(* IEC 61131-3 sources: MongoMation/docs, 1 file *)

(* ---- probe-sorting-by-height-basic.st ---- *)
(* I/O probe for scene sorting-by-height-basic (Sorting by Height (Basic)). Generated by scripts/gen-probe.ts. *)
PROGRAM io_probe
  VAR
    I0 AT %QX12.4 : BOOL; (* High sensor *)
    I1 AT %QX12.5 : BOOL; (* Low sensor *)
    I2 AT %QX12.6 : BOOL; (* Pallet sensor *)
    I3 AT %QX12.7 : BOOL; (* Loaded *)
    I4 AT %QX13.0 : BOOL; (* At left entry *)
    I5 AT %QX13.1 : BOOL; (* At left exit *)
    I6 AT %QX13.2 : BOOL; (* At right entry *)
    I7 AT %QX13.3 : BOOL; (* At right exit *)
    I8 AT %QX13.4 : BOOL; (* Start *)
    I9 AT %QX13.5 : BOOL; (* Reset *)
    I10 AT %QX13.6 : BOOL; (* Stop *)
    I11 AT %QX13.7 : BOOL; (* Emergency stop *)
    I12 AT %QX14.0 : BOOL; (* Auto *)
    Q0 AT %QX0.0 : BOOL; (* Conveyor entry *)
    Q1 AT %QX0.1 : BOOL; (* Load *)
    Q2 AT %QX0.2 : BOOL; (* Unload *)
    Q3 AT %QX0.3 : BOOL; (* Transf. left *)
    Q4 AT %QX0.4 : BOOL; (* Transf. right *)
    Q5 AT %QX0.5 : BOOL; (* Conveyor left *)
    Q6 AT %QX0.6 : BOOL; (* Conveyor right *)
    Q7 AT %QX0.7 : BOOL; (* Start light *)
    Q8 AT %QX1.0 : BOOL; (* Reset light *)
    Q9 AT %QX1.1 : BOOL; (* Stop light *)
  END_VAR
  VAR
    Tick : TON;
    Phase : INT := 0;
    InputsSeen : INT := 0;
  END_VAR
  Tick(IN := NOT Tick.Q, PT := T#1000ms);
  IF Tick.Q THEN
    Phase := Phase + 1;
    IF Phase >= 10 THEN
      Phase := 0;
    END_IF;
  END_IF;
  Q0 := (Phase = 0); (* Conveyor entry *)
  Q1 := (Phase = 1); (* Load *)
  Q2 := (Phase = 2); (* Unload *)
  Q3 := (Phase = 3); (* Transf. left *)
  Q4 := (Phase = 4); (* Transf. right *)
  Q5 := (Phase = 5); (* Conveyor left *)
  Q6 := (Phase = 6); (* Conveyor right *)
  Q7 := (Phase = 7); (* Start light *)
  Q8 := (Phase = 8); (* Reset light *)
  Q9 := (Phase = 9); (* Stop light *)
  InputsSeen := 0;
  IF I0 THEN InputsSeen := InputsSeen + 1; END_IF;
  IF I1 THEN InputsSeen := InputsSeen + 1; END_IF;
  IF I2 THEN InputsSeen := InputsSeen + 1; END_IF;
  IF I3 THEN InputsSeen := InputsSeen + 1; END_IF;
  IF I4 THEN InputsSeen := InputsSeen + 1; END_IF;
  IF I5 THEN InputsSeen := InputsSeen + 1; END_IF;
  IF I6 THEN InputsSeen := InputsSeen + 1; END_IF;
  IF I7 THEN InputsSeen := InputsSeen + 1; END_IF;
  IF I8 THEN InputsSeen := InputsSeen + 1; END_IF;
  IF I9 THEN InputsSeen := InputsSeen + 1; END_IF;
  IF I10 THEN InputsSeen := InputsSeen + 1; END_IF;
  IF I11 THEN InputsSeen := InputsSeen + 1; END_IF;
  IF I12 THEN InputsSeen := InputsSeen + 1; END_IF;
END_PROGRAM

CONFIGURATION Config0
  RESOURCE Res0 ON PLC
    TASK task0(INTERVAL := T#20ms, PRIORITY := 0);
    PROGRAM instance0 WITH task0 : io_probe;
  END_RESOURCE
END_CONFIGURATION
